// TIA Portal V21 export
// export: Created 2026-11-11T00:47:34.8930569Z, ExportSetting WithDefaults, DisplayName Totally Integrated Automation Portal, DisplayVersion V21 Update 3, DisplayName STEP 7 Professional, DisplayVersion V21 Update 3, DisplayName STEP 7 Safety, DisplayVersion V21, DisplayName Tech WebApplication, DisplayVersion V21, DisplayName WinCC Basic/Comfort/Advanced, DisplayVersion V21 Update 3, DisplayName WinCC Unified, DisplayVersion V21 Update 3
FUNCTION_BLOCK "FB_Fbd_ex132"   // FB142, FBD
{ S7_Optimized_Access := 'TRUE' }
VERSION : 0.1
// stored: AutoNumber true, IsIECCheckEnabled false, IsRetainMemResEnabled false, MemoryReserve 100, SetENOAutomatically false, UDAEnableTagReadback false
   VAR_INPUT
      v_laddr : HW_ANY;
      v_mode : UInt;
   END_VAR
   VAR_OUTPUT
      v_ret_val : Int;
   END_VAR
   VAR_IN_OUT
      v_diagevent : DiagnosticDetail;
   END_VAR
BEGIN

REGION Network 1: GEN_DIAG - Generate diagnostics information
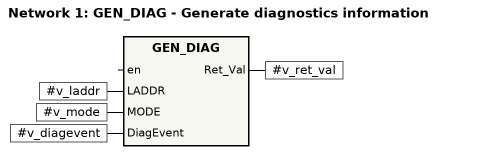
   #v_ret_val := GEN_DIAG(LADDR := #v_laddr, MODE := #v_mode, DiagEvent := #v_diagevent);
END_REGION
END_FUNCTION_BLOCK
